TYPE ST_AutomaticExtractionHandlerTest :
STRUCT
	automaticExtractionStateMachine : ST_AutomaticExtractionStateMachineTest;
END_STRUCT
END_TYPE

(* stored: Version 1.1.0.1, ProductVersion 3.1.4024.9
   DUT ST_AutomaticExtractionHandlerTest: Id {e42ec552-f74d-4d23-8cdc-569a909abd1c} *)
